Fanuc KAREL source: KX00010.KL

PROGRAM KX00010
%NOLOCKGROUP
VAR
  I: INTEGER
  J: INTEGER
  B: BOOLEAN
  F: FILE
  S: STRING[80]
  P: XYZWPR
BEGIN
  PAUSE
END KX00010
